// Mitsubishi GX Works2 project: 261019_적산 타이머 실습_타이머 추가 응용2   PLC: Q03UDV

PROGRAM MAIN
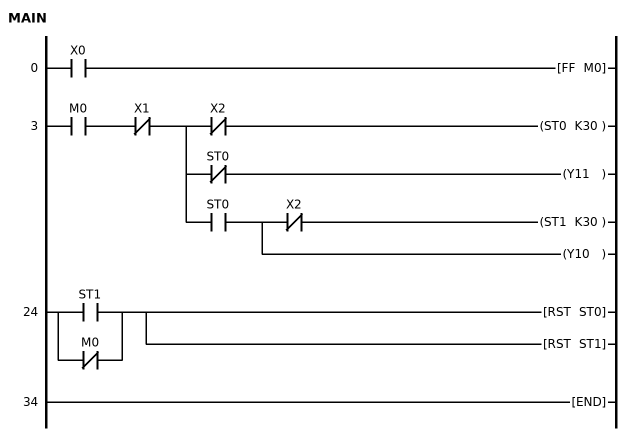
0     LD      X0
      FF      M0
3     LD      M0
      ANI     X1
      MPS
      ANI     X2
      OUT     ST0 K30
      MRD
      ANI     ST0
      OUT     Y11
      MPP
      AND     ST0
      MPS
      ANI     X2
      OUT     ST1 K30
      MPP
      OUT     Y10
24    LD      ST1
      ORI     M0
      RST     ST0
      RST     ST1
34    END
END_PROGRAM
